// TIA Portal V21 export
// export: Created 2026-11-10T19:11:40.8115974Z, ExportSetting WithDefaults, DisplayName Totally Integrated Automation Portal, DisplayVersion V21 Update 3, DisplayName STEP 7 Professional, DisplayVersion V21 Update 3, DisplayName STEP 7 Safety, DisplayVersion V21, DisplayName Tech WebApplication, DisplayVersion V21, DisplayName WinCC Basic/Comfort/Advanced, DisplayVersion V21 Update 3, DisplayName WinCC Unified, DisplayVersion V21 Update 3
DATA_BLOCK "DB_RALRM_SFB"   // DB50
// stored: AutoNumber true, DBAccessibleFromOPCUA true, DBAccessibleFromWebserver true, InstanceOfName RALRM_SFB, OfSystemLibElement RALRM, OfSystemLibVersion 1.0
"RALRM_SFB"
   // VAR_INPUT
   //    MODE : Int;
   //    F_ID : HW_IO;
   //    MLEN : UInt;
   // END_VAR
   // VAR_OUTPUT
   //    NEW : Bool;
   //    STATUS : DWord;
   //    ID : HW_IO;
   //    LEN : UInt;
   // END_VAR
   // VAR_IN_OUT
   //    TINFO : Variant;
   //    AINFO : Variant;
   // END_VAR
BEGIN
END_DATA_BLOCK
